TYPE ST_PositionProcess :
STRUCT
	lrProcessPosition						:LREAL;											(* Process position [mm] *)
	unProcessVelo						:UINT;											(* Process force [%] *)
	unProcessRamp						:UINT;											(* Process ramp [s] *)
	unProcessTime						:UINT;											(* Process time [s]  *)
	arunDuration							:ARRAY[1..2] OF UINT;								(* Duration [s] *)
END_STRUCT
END_TYPE

(* stored: Version 1.1.0.1, ProductVersion 3.1.4024.15
   DUT ST_PositionProcess: Id {9f497c85-f4ea-4a5d-b4f3-b24858a1faa4} *)
